Universal Robots PolyScope program: Sub_AMR_MiR_V3.urp

Program Sub_AMR_MiR_V3 (installation=default directory=/programs/03 Sub Routines createdIn=5.11.11 lastSavedIn=5.23.0 robotSerialNumber=20245590049)
Calibrated DH parameters: a=[0.000139, -0.197451, -0.383992, -0.000109, 0.000038, 0]; d=[0.162494, 274.063354, -251.846761, -22.083037, 0.099612, 0.099364]; alpha=[1.570089, 0.001374, 0.003592, 1.570222, -1.570187, 0]; deltaTheta=[0, 1.08787, 5.400214, -0.204909, 0.000001, 0]
InitVariablesNode variables(variable(name=AMR_Position, expression=struct(position_identifier=0, x1=0, x2=0, y1=0, y2=0, theta1=0, theta2=0)), variable(name=CAM_Pose, expression=p[0,0,0,0,0,0]), variable(name=CAM_Relation, expression=""), variable(name=CMD_Abort, expression=False), variable(name=CMD_Clear, expression=False), variable(name=CMD_Reset, expression=False), variable(name=CMD_Start, expression=False), variable(name=CMD_Suspend, expression=False), variable(name=CMD_Unhold, expression=False), variable(name=CMD_Unsuspend, expression=False), variable(name=CNT_Rack_Output, expression=0), variable(name=FNC_Freedrive, expression=False), variable(name=PRC_TubCounter, expression=0), variable(name=STP, expression=0), variable(name=TMR_Barcode, expression=0), variable(name=easyPickCount_4, expression=0), variable(name=easyPickCount_7, expression=0), variable(name=easyPickNoObj_4, expression=0), variable(name=easyPickNoObj_7, expression=0), variable(name=easyPickParts_4, expression=0), variable(name=easyPickParts_7, expression=0))
BeforeStart
  Folder Manual
    SafeHome (positionOptionType=SPEED_AND_ACCELERATION speed=1.047198 acceleration=1.396263 nextMotionTime=2)
    STATE :=  (valueSource=Operator message=state valueType=Integer)
    If STATE≟6
      Action :=  (valueSource=Operator message=what valueType=Integer)
      If Action≟52
        AMR_PosTarget :=  (valueSource=Operator message=target valueType=Integer)
Robot Program (runOnlyOnce=true)
  Folder PreSettings [hidden by the author, left out]
  '=========='
  Switch expression=STATE
    Case (caseValue=1)
      Folder stopping
        If T2O_Done≟1 and O2T_Acknowledge≟0
          Set ExpressionOutput pin=O2T_Acknowledge; expression=1
        Set DigitalOutput pin=MiR_CMD_Stop; digitalValue=1
        Script: AMR_Position.position_identifier = 0
        AMR_Done := True
    Case (caseValue=2)
      Folder stopped
        If MiR_State≠3 and MiR_State≠5
          Set DigitalOutput pin=MiR_CMD_Stop; digitalValue=0
    Case (caseValue=3)
      Folder resetting [hidden by the author, left out]
    Case (caseValue=5)
      Folder starting
        If MiR_State≟4
          Set DigitalOutput pin=MiR_CMD_Start; digitalValue=1
          Wait Condition expression=MiR_State≠4
          Set DigitalOutput pin=MiR_CMD_Start; digitalValue=0
          AMR_Done := True
        ElseIf MiR_State≟10
          'MiR in protective stop. Wait'
          AMR_Done := True
        ElseIf MiR_State≟3
          AMR_Done := True
    Case (caseValue=6)
      Folder execute
        AMR_AtTarget := (AMR_PosActual≟AMR_PosTarget)
        Switch expression=AMR_Step
          Case (caseValue=0)
            If not AMR_AtTarget
              AMR_Step := 1
            Else 
              AMR_Done := True
          Case (caseValue=1)
            Folder general Settings [hidden by the author, left out]
            Folder check for error
              If OBJ_Picked and MiR_State≟10
                Folder Error
                  Script: set_error(ERROR_ROBOT_ARM_NOT_IN_HOME_POSE)
                Action := 0
              ElseIf not found_in_list(AMR_PosTarget, AMR_TargetList)
                Folder Error
                  Script: set_error(ERROR_UNKNOWN_POSE)
                Action := 0
            If MiR_State≟3
              Set DigitalOutput pin=MiR_CMD_Start; digitalValue=0
              Switch expression=Action
                Case (caseValue=51)
                  Folder Charge
                    'trigger the charging mission'
                    'target pos is predefined'
                    Set ExpressionOutput pin=O2T_Footprint; expression=0
                    Set ExpressionOutput pin=O2T_Action; expression=1
                  If MiR_Mis_Queue≟0
                    Set DigitalOutput pin=O2T_Mis_Charge; digitalValue=1
                    Wait Condition expression=MiR_Mis_Queue≥1
                    Set DigitalOutput pin=O2T_Mis_Charge; digitalValue=0
                Case (caseValue=52)
                  Folder Navigate
                    'trigger the standard missoin'
                    Set ExpressionOutput pin=O2T_Footprint; expression=AMR_FootprintID
                    Set ExpressionOutput pin=O2T_Target_Pos; expression=AMR_PosTarget
                    Set ExpressionOutput pin=O2T_Action; expression=2
                  If MiR_Mis_Queue≟0
                    Set DigitalOutput pin=O2T_Mis_Main; digitalValue=1
                    Wait Condition expression=MiR_Mis_Queue≥1
                    Set DigitalOutput pin=O2T_Mis_Main; digitalValue=0
            ElseIf MiR_State≟4
              Set DigitalOutput pin=MiR_CMD_Start; digitalValue=1
            ElseIf MiR_State≟5
              AMR_Step := 2
            ElseIf MiR_State≟10
              'AMR still in safeguard stop'
          Case (caseValue=2)
            Folder acknowledge handshake
              If T2O_Done≟1 and O2T_Acknowledge≟0
                Set ExpressionOutput pin=O2T_Acknowledge; expression=1
              ElseIf T2O_Done≟0 and O2T_Acknowledge≟1
                Set ExpressionOutput pin=O2T_Acknowledge; expression=0
                AMR_AtTarget := (AMR_PosActual≟AMR_PosTarget)
                AMR_Done := True
        Folder translate errors [hidden by the author, left out]
    Case (caseValue=7)
      Folder completing [hidden by the author, left out]
    Case (caseValue=9)
      Folder holding [hidden by the author, left out]
    Case (caseValue=11)
      Folder unholding [hidden by the author, left out]
    Case (caseValue=12)
      Folder suspending [hidden by the author, left out]
    Case (caseValue=14)
      Folder unsuspending [hidden by the author, left out]
    Case (caseValue=15)
      Folder aborting [hidden by the author, left out]
    Case (caseValue=17)
      Folder clearing [hidden by the author, left out]
  '=========='
  Folder PostSettings [hidden by the author, left out]
